(* IEC 61131-3 sources: kns-port-domestic/upstream/kns-pump-station/src/POUs/Generated/PRG_Devices, 2 files *)

(* ---- PRG_Devices.decl.st ---- *)
// AUTO-GENERATED by iolistgen 0.2.0 — не редактировать; источник: 03_io_list.csv
// SHA-256 перечня 06336d13c4b2; генератор st-codesys
// Назначение: вызовы устройств plc-process-lib по перечню сигналов: входы из GVL_IO, выходы в GVL_IO, команды GVL_Hmi,
// Cfg и Retain — GVL_Persist (контракт plc-process-lib, разделы 1 и 20). Входы автоматики (xAutoRun, xAutoOpen,
// wInterlock, wPermit…, rSpeedSpAuto_pct, rPosSpAuto_pct) пишет логика станции до вызова PRG_Devices
// Автор:      iolistgen (генератор по перечню сигналов); перечень 03_io_list.csv
// Версия:     iolistgen 0.2.0
// Документ:   docs/03_io_list.md
PROGRAM PRG_Devices
VAR
END_VAR

(* ---- PRG_Devices.impl.st ---- *)
// AUTO-GENERATED by iolistgen 0.2.0 — не редактировать; источник: 03_io_list.csv
// SHA-256 перечня 06336d13c4b2; генератор st-codesys
// Порядок: устройства, на которые ссылаются link_power и link_fb (ES301), вызываются раньше ссылающихся; дальше — по
// dev_no.

// КНС-1 (перекрытие шаблона iolistgen, docs/DESIGN.md, раздел 4.6): входы GVL_IO недействительны, пока в
// имитации модель не опубликовала их ни разу (PlantModelTask ниже MainTask по приоритету: первый цикл MainTask
// видит нули). Первый вызов устройств — подхват и начальные значения DI — только по действительным входам
IF NOT GVL_Sim.xIoReady THEN
    RETURN;
END_IF

// Приёмник событий тревог библиотеки: присваивается каждый цикл до вызова устройств (контракт 5.3)
PL.GVL_Lib.itfAlarmSink := GVL_Log.fbEventLog;

// Команда HMI «Применить уставки проекта» (контракт 18.3, правило 2): Retain устройств не меняется
IF GVL_Hmi.xApplyProjectCfg THEN
    GVL_Hmi.xApplyProjectCfg := FALSE;
    PRG_ApplyProjectCfg();
END_IF

// --- dev_no 301: ES301 — Напряжение на вводе в норме (реле контроля фаз) (DigitalInput) ---
GVL_Devices.fbES301(
    xIn           := GVL_IO.xES301,
    xChannelFault := FALSE,  // нет строки CHF
    itfTime       := GVL_Time.fbClockMain,  // источник времени
    stCmd         := GVL_Hmi.stES301Cmd,
    stCfg         := GVL_Persist.stES301Cfg);

// --- dev_no 11: P101 — Насос Н1 (MotorVfd) ---
// ПЧ: xCommOk, xVfd*, rSpeedAct_pct и rSpeedRef_pct — через адаптер приложения (GVL_IO.xP101_…)
// без входа ФБ (AUX, код приложения): GVL_IO.uiP101_FCODE — Насос Н1: код последней аварии ПЧ (читает адаптер ПЧ)
GVL_Devices.fbP101(
    xFbRun        := GVL_IO.xP101_RFB,
    xExtFault     := GVL_IO.xP101_FLT,
    xLocal        := GVL_IO.xHS114,
    xPowerOk      := GVL_Devices.fbES301.xValue,  // link_power
    xCommOk       := GVL_IO.xP101_CommOk,
    xVfdRunning   := GVL_IO.xP101_VfdRun,
    xVfdReady     := GVL_IO.xP101_VfdReady,
    xVfdFault     := GVL_IO.xP101_VfdFault,
    rSpeedAct_pct := GVL_IO.rP101_SpeedAct_pct,
    itfTime       := GVL_Time.fbClockMain,  // источник времени
    stCmd         := GVL_Hmi.stP101Cmd,
    stCfg         := GVL_Persist.stP101Cfg,
    stRetain      := GVL_Persist.stP101Retain);
GVL_IO.xP101_RUN          := GVL_Devices.fbP101.xQRun;
GVL_IO.xP101_VfdQRun      := GVL_Devices.fbP101.xQRun;
GVL_IO.xP101_VfdQReset    := GVL_Devices.fbP101.xQReset;
GVL_IO.rP101_SpeedRef_pct := GVL_Devices.fbP101.rSpeedRef_pct;

// --- dev_no 12: P102 — Насос Н2 (MotorVfd) ---
// ПЧ: xCommOk, xVfd*, rSpeedAct_pct и rSpeedRef_pct — через адаптер приложения (GVL_IO.xP102_…)
// без входа ФБ (AUX, код приложения): GVL_IO.uiP102_FCODE — Насос Н2: код последней аварии ПЧ (читает адаптер ПЧ)
GVL_Devices.fbP102(
    xFbRun        := GVL_IO.xP102_RFB,
    xExtFault     := GVL_IO.xP102_FLT,
    xLocal        := GVL_IO.xHS124,
    xPowerOk      := GVL_Devices.fbES301.xValue,  // link_power
    xCommOk       := GVL_IO.xP102_CommOk,
    xVfdRunning   := GVL_IO.xP102_VfdRun,
    xVfdReady     := GVL_IO.xP102_VfdReady,
    xVfdFault     := GVL_IO.xP102_VfdFault,
    rSpeedAct_pct := GVL_IO.rP102_SpeedAct_pct,
    itfTime       := GVL_Time.fbClockMain,  // источник времени
    stCmd         := GVL_Hmi.stP102Cmd,
    stCfg         := GVL_Persist.stP102Cfg,
    stRetain      := GVL_Persist.stP102Retain);
GVL_IO.xP102_RUN          := GVL_Devices.fbP102.xQRun;
GVL_IO.xP102_VfdQRun      := GVL_Devices.fbP102.xQRun;
GVL_IO.xP102_VfdQReset    := GVL_Devices.fbP102.xQReset;
GVL_IO.rP102_SpeedRef_pct := GVL_Devices.fbP102.rSpeedRef_pct;

// --- dev_no 13: P103 — Насос Н3 (MotorVfd) ---
// ПЧ: xCommOk, xVfd*, rSpeedAct_pct и rSpeedRef_pct — через адаптер приложения (GVL_IO.xP103_…)
// без входа ФБ (AUX, код приложения): GVL_IO.uiP103_FCODE — Насос Н3: код последней аварии ПЧ (читает адаптер ПЧ)
GVL_Devices.fbP103(
    xFbRun        := GVL_IO.xP103_RFB,
    xExtFault     := GVL_IO.xP103_FLT,
    xLocal        := GVL_IO.xHS134,
    xPowerOk      := GVL_Devices.fbES301.xValue,  // link_power
    xCommOk       := GVL_IO.xP103_CommOk,
    xVfdRunning   := GVL_IO.xP103_VfdRun,
    xVfdReady     := GVL_IO.xP103_VfdReady,
    xVfdFault     := GVL_IO.xP103_VfdFault,
    rSpeedAct_pct := GVL_IO.rP103_SpeedAct_pct,
    itfTime       := GVL_Time.fbClockMain,  // источник времени
    stCmd         := GVL_Hmi.stP103Cmd,
    stCfg         := GVL_Persist.stP103Cfg,
    stRetain      := GVL_Persist.stP103Retain);
GVL_IO.xP103_RUN          := GVL_Devices.fbP103.xQRun;
GVL_IO.xP103_VfdQRun      := GVL_Devices.fbP103.xQRun;
GVL_IO.xP103_VfdQReset    := GVL_Devices.fbP103.xQReset;
GVL_IO.rP103_SpeedRef_pct := GVL_Devices.fbP103.rSpeedRef_pct;

// --- dev_no 14: V1 — Вытяжной вентилятор В1 павильона (Motor) ---
GVL_Devices.fbV1(
    xFbRun    := GVL_IO.xV1_RFB,
    xExtFault := GVL_IO.xV1_FLT,
    xPowerOk  := GVL_Devices.fbES301.xValue,  // link_power
    itfTime   := GVL_Time.fbClockMain,  // источник времени
    stCmd     := GVL_Hmi.stV1Cmd,
    stCfg     := GVL_Persist.stV1Cfg,
    stRetain  := GVL_Persist.stV1Retain);
GVL_IO.xV1_RUN := GVL_Devices.fbV1.xQRun;

// --- dev_no 101: LT101 — Уровень в приёмном резервуаре (AnalogInput) ---
GVL_Devices.fbLT101(
    rIn           := GVL_IO.rLT101_mA,
    xChannelFault := FALSE,  // нет строки CHF
    itfTime       := GVL_Time.fbClockMain,  // источник времени
    stCmd         := GVL_Hmi.stLT101Cmd,
    stCfg         := GVL_Persist.stLT101Cfg);

// --- dev_no 102: LS102 — Поплавок «аварийно высокий уровень» (H, 4,2 м) (DigitalInput) ---
GVL_Devices.fbLS102(
    xIn           := GVL_IO.xLS102,
    xChannelFault := FALSE,  // нет строки CHF
    itfTime       := GVL_Time.fbClockMain,  // источник времени
    stCmd         := GVL_Hmi.stLS102Cmd,
    stCfg         := GVL_Persist.stLS102Cfg);

// --- dev_no 103: LS103 — Поплавок «сухой ход» (L, 0,4 м) (DigitalInput) ---
GVL_Devices.fbLS103(
    xIn           := GVL_IO.xLS103,
    xChannelFault := FALSE,  // нет строки CHF
    itfTime       := GVL_Time.fbClockMain,  // источник времени
    stCmd         := GVL_Hmi.stLS103Cmd,
    stCfg         := GVL_Persist.stLS103Cfg);

// --- dev_no 111: IT111 — Насос Н1: ток двигателя (измеряет ПЧ) (AnalogInput) ---
GVL_Devices.fbIT111(
    rIn           := UINT_TO_REAL(GVL_IO.uiIT111),
    xChannelFault := NOT GVL_IO.xMbOk_RS485_1_S1,  // нет строки CHF: обмен со слейвом
    itfTime       := GVL_Time.fbClockMain,  // источник времени
    stCmd         := GVL_Hmi.stIT111Cmd,
    stCfg         := GVL_Persist.stIT111Cfg);

// --- dev_no 112: TS112 — Насос Н1: перегрев обмотки (термовыключатели, реле защиты насоса) (DigitalInput) ---
GVL_Devices.fbTS112(
    xIn           := GVL_IO.xTS112,
    xChannelFault := FALSE,  // нет строки CHF
    itfTime       := GVL_Time.fbClockMain,  // источник времени
    stCmd         := GVL_Hmi.stTS112Cmd,
    stCfg         := GVL_Persist.stTS112Cfg);

// --- dev_no 113: MS113 — Насос Н1: протечка в камеру статора (датчик влажности, реле защиты насоса) (DigitalInput) ---
GVL_Devices.fbMS113(
    xIn           := GVL_IO.xMS113,
    xChannelFault := FALSE,  // нет строки CHF
    itfTime       := GVL_Time.fbClockMain,  // источник времени
    stCmd         := GVL_Hmi.stMS113Cmd,
    stCfg         := GVL_Persist.stMS113Cfg);

// --- dev_no 121: IT121 — Насос Н2: ток двигателя (измеряет ПЧ) (AnalogInput) ---
GVL_Devices.fbIT121(
    rIn           := UINT_TO_REAL(GVL_IO.uiIT121),
    xChannelFault := NOT GVL_IO.xMbOk_RS485_1_S2,  // нет строки CHF: обмен со слейвом
    itfTime       := GVL_Time.fbClockMain,  // источник времени
    stCmd         := GVL_Hmi.stIT121Cmd,
    stCfg         := GVL_Persist.stIT121Cfg);

// --- dev_no 122: TS122 — Насос Н2: перегрев обмотки (термовыключатели, реле защиты насоса) (DigitalInput) ---
GVL_Devices.fbTS122(
    xIn           := GVL_IO.xTS122,
    xChannelFault := FALSE,  // нет строки CHF
    itfTime       := GVL_Time.fbClockMain,  // источник времени
    stCmd         := GVL_Hmi.stTS122Cmd,
    stCfg         := GVL_Persist.stTS122Cfg);

// --- dev_no 123: MS123 — Насос Н2: протечка в камеру статора (датчик влажности, реле защиты насоса) (DigitalInput) ---
GVL_Devices.fbMS123(
    xIn           := GVL_IO.xMS123,
    xChannelFault := FALSE,  // нет строки CHF
    itfTime       := GVL_Time.fbClockMain,  // источник времени
    stCmd         := GVL_Hmi.stMS123Cmd,
    stCfg         := GVL_Persist.stMS123Cfg);

// --- dev_no 131: IT131 — Насос Н3: ток двигателя (измеряет ПЧ) (AnalogInput) ---
GVL_Devices.fbIT131(
    rIn           := UINT_TO_REAL(GVL_IO.uiIT131),
    xChannelFault := NOT GVL_IO.xMbOk_RS485_1_S3,  // нет строки CHF: обмен со слейвом
    itfTime       := GVL_Time.fbClockMain,  // источник времени
    stCmd         := GVL_Hmi.stIT131Cmd,
    stCfg         := GVL_Persist.stIT131Cfg);

// --- dev_no 132: TS132 — Насос Н3: перегрев обмотки (термовыключатели, реле защиты насоса) (DigitalInput) ---
GVL_Devices.fbTS132(
    xIn           := GVL_IO.xTS132,
    xChannelFault := FALSE,  // нет строки CHF
    itfTime       := GVL_Time.fbClockMain,  // источник времени
    stCmd         := GVL_Hmi.stTS132Cmd,
    stCfg         := GVL_Persist.stTS132Cfg);

// --- dev_no 133: MS133 — Насос Н3: протечка в камеру статора (датчик влажности, реле защиты насоса) (DigitalInput) ---
GVL_Devices.fbMS133(
    xIn           := GVL_IO.xMS133,
    xChannelFault := FALSE,  // нет строки CHF
    itfTime       := GVL_Time.fbClockMain,  // источник времени
    stCmd         := GVL_Hmi.stMS133Cmd,
    stCfg         := GVL_Persist.stMS133Cfg);

// --- dev_no 201: PT201 — Давление в напорном коллекторе (AnalogInput) ---
GVL_Devices.fbPT201(
    rIn           := GVL_IO.rPT201_mA,
    xChannelFault := FALSE,  // нет строки CHF
    itfTime       := GVL_Time.fbClockMain,  // источник времени
    stCmd         := GVL_Hmi.stPT201Cmd,
    stCfg         := GVL_Persist.stPT201Cfg);

// --- dev_no 202: FT202 — Расход в напорном коллекторе (AnalogInput) ---
GVL_Devices.fbFT202(
    rIn           := GVL_IO.rFT202_mA,
    xChannelFault := FALSE,  // нет строки CHF
    itfTime       := GVL_Time.fbClockMain,  // источник времени
    stCmd         := GVL_Hmi.stFT202Cmd,
    stCfg         := GVL_Persist.stFT202Cfg);

// --- dev_no 203: LS203 — Затопление камеры задвижек (DigitalInput) ---
GVL_Devices.fbLS203(
    xIn           := GVL_IO.xLS203,
    xChannelFault := FALSE,  // нет строки CHF
    itfTime       := GVL_Time.fbClockMain,  // источник времени
    stCmd         := GVL_Hmi.stLS203Cmd,
    stCfg         := GVL_Persist.stLS203Cfg);

// --- dev_no 302: YS302 — ИБП шкафа управления: работа от батарей (DigitalInput) ---
GVL_Devices.fbYS302(
    xIn           := GVL_IO.xYS302,
    xChannelFault := FALSE,  // нет строки CHF
    itfTime       := GVL_Time.fbClockMain,  // источник времени
    stCmd         := GVL_Hmi.stYS302Cmd,
    stCfg         := GVL_Persist.stYS302Cfg);

// --- dev_no 303: YS303 — ИБП шкафа управления: неисправность или разряд батарей (DigitalInput) ---
GVL_Devices.fbYS303(
    xIn           := GVL_IO.xYS303,
    xChannelFault := FALSE,  // нет строки CHF
    itfTime       := GVL_Time.fbClockMain,  // источник времени
    stCmd         := GVL_Hmi.stYS303Cmd,
    stCfg         := GVL_Persist.stYS303Cfg);

// --- dev_no 401: AT401 — Концентрация сероводорода H₂S в павильоне (AnalogInput) ---
GVL_Devices.fbAT401(
    rIn           := GVL_IO.rAT401_mA,
    xChannelFault := FALSE,  // нет строки CHF
    itfTime       := GVL_Time.fbClockMain,  // источник времени
    stCmd         := GVL_Hmi.stAT401Cmd,
    stCfg         := GVL_Persist.stAT401Cfg);

// --- dev_no 402: AT402 — Концентрация метана CH₄ в павильоне (AnalogInput) ---
GVL_Devices.fbAT402(
    rIn           := GVL_IO.rAT402_mA,
    xChannelFault := FALSE,  // нет строки CHF
    itfTime       := GVL_Time.fbClockMain,  // источник времени
    stCmd         := GVL_Hmi.stAT402Cmd,
    stCfg         := GVL_Persist.stAT402Cfg);

// --- dev_no 403: TT403 — Температура воздуха в павильоне (AnalogInput) ---
GVL_Devices.fbTT403(
    rIn           := GVL_IO.rTT403,
    xChannelFault := NOT GVL_IO.xMbOk_RS485_2_S10,  // нет строки CHF: обмен со слейвом
    itfTime       := GVL_Time.fbClockMain,  // источник времени
    stCmd         := GVL_Hmi.stTT403Cmd,
    stCfg         := GVL_Persist.stTT403Cfg);

// --- dev_no 404: ZS404 — Дверь павильона открыта (DigitalInput) ---
GVL_Devices.fbZS404(
    xIn           := GVL_IO.xZS404,
    xChannelFault := FALSE,  // нет строки CHF
    itfTime       := GVL_Time.fbClockMain,  // источник времени
    stCmd         := GVL_Hmi.stZS404Cmd,
    stCfg         := GVL_Persist.stZS404Cfg);

// --- dev_no 405: YS405 — Пожар (сигнал прибора пожарной сигнализации) (DigitalInput) ---
GVL_Devices.fbYS405(
    xIn           := GVL_IO.xYS405,
    xChannelFault := FALSE,  // нет строки CHF
    itfTime       := GVL_Time.fbClockMain,  // источник времени
    stCmd         := GVL_Hmi.stYS405Cmd,
    stCfg         := GVL_Persist.stYS405Cfg);

// --- dev_no 501: HS501 — Кнопка «Сброс аварий» на двери шкафа управления (DigitalInput) ---
GVL_Devices.fbHS501(
    xIn           := GVL_IO.xHS501,
    xChannelFault := FALSE,  // нет строки CHF
    itfTime       := GVL_Time.fbClockMain,  // источник времени
    stCmd         := GVL_Hmi.stHS501Cmd,
    stCfg         := GVL_Persist.stHS501Cfg);

// --- dev_no 502: HS502 — Кнопка «Отключить звук» на двери шкафа управления (DigitalInput) ---
GVL_Devices.fbHS502(
    xIn           := GVL_IO.xHS502,
    xChannelFault := FALSE,  // нет строки CHF
    itfTime       := GVL_Time.fbClockMain,  // источник времени
    stCmd         := GVL_Hmi.stHS502Cmd,
    stCfg         := GVL_Persist.stHS502Cfg);
